Yaskawa INFORM job: SETPROG.JBI

/JOB
//NAME SETPROG
//POS
///NPOS 7,0,0,0,0,0
///TOOL 9
///POSTYPE PULSE
///PULSE
C00000=0,-19456,25243,0,27307,0
C00001=0,-19456,25243,0,27307,0
C00002=0,-19456,25243,0,27307,0
C00003=0,-19456,25243,0,27307,0
C00004=36064,-19456,25243,0,27307,0
C00005=36064,-19456,25243,0,27307,0
C00006=54096,-38912,50486,64027,-40960,-56268
//INST
<volatile>
///COMM Generated using RoboDK
///ATTR SC,RW
///GROUP1 RB1
NOP
'Program generated by RoboDK v
'6.0.7 for Yaskawa Motoman DX1
'350D on XX/XX/XXXX 18:00:00
'Using nominal kinematics.
'Using Frame S (targets wrt ba
'se):
'1234.6,-98.8,50.5,0.0,0.0,30.
'0
'Tool Tool S should be close t
'o:
'10.0,20.0,150.0,0.0,0.0,0.0
MOVJ C00000 VJ=50.00
MOVL C00001 V=100.0
MOVC C00002 V=100.0
MOVC C00003 V=100.0
MOVC C00004 V=100.0
MOVJ C00005 VJ=50.00
TIMER T=0.25
MOVJ C00006 VJ=50.00
END
